ABB RobotStudio station: FrezaEGM_20261120-133356.rsstn

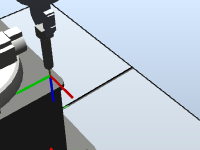
Station FrezaEGM (saved by RobotStudio 6.8.8307.1040)
Controller FrezaEGM, task T_ROB1: task frame (RAPID world) sits at (0, 0, 520) mm in the station
Controller FrezaEGM
  mechanical unit ROB_1: IRB1600_10_145__01, 6 joints, base frame (0, 0, 0) mm
Layout (positions relative to the parent item):
  - IRB1600_10_145__01 [mechanism, from Robots\IRB1600_10_145_G_01.rslib] at (0, 0, 520) mm; joint values [0, 0.0714, 0.3396, 0, 1.1598, 3.1416] (rad or m)
  - подставка [part, from Libraries\подставка.rslib]
  - toolPencil [mechanism, from Libraries\toolPencil.rslib] at (750, 0, 1400) mm, rotated rx -180 ry 0 rz 0 deg
Attachment: toolPencil is attached to IRB1600_10_145__01 / Link6
Targets, tools, work objects and paths stored in the station, written as RAPID:
! task T_ROB1
MODULE ModuleEGM
  LOCAL CONST robtarget home:=[[750,0,300],[0,0,1,0],[0,0,0,0],[9E+09,0,0,9E+09,9E+09,9E+09]];
  PROC main()
    MoveJ home,v100,fine,tool0;
  ENDPROC
ENDMODULE

! task T_ROB1
MODULE CalibData
  PERS tooldata toolPencil:=[TRUE,[[0,0,280],[1,0,0,0]],[1,[0,0,1],[1,0,0,0],0,0,0]];
ENDMODULE

